// TIA Portal V21 export
// export: Created 2026-11-10T07:35:08.0372515Z, ExportSetting WithDefaults, DisplayName Totally Integrated Automation Portal, DisplayVersion V21 Update 3, DisplayName STEP 7 Professional, DisplayVersion V21 Update 3, DisplayName STEP 7 Safety, DisplayVersion V21, DisplayName Tech WebApplication, DisplayVersion V21, DisplayName WinCC Basic/Comfort/Advanced, DisplayVersion V21 Update 3, DisplayName WinCC Unified, DisplayVersion V21 Update 3
FUNCTION_BLOCK "FB_Lad_ex063"   // FB98, LAD
{ S7_Optimized_Access := 'TRUE' }
VERSION : 0.1
// stored: AutoNumber true, IsIECCheckEnabled false, IsRetainMemResEnabled false, MemoryReserve 100, SetENOAutomatically false, UDAEnableTagReadback false
   VAR_INPUT
      v_mode : Int;
      v_f_id : HW_SUBMODULE;
      v_code1 : Byte;
      v_code2 : Byte;
      v_len : UInt;
   END_VAR
   VAR_OUTPUT
      v_new : Bool;
      v_status : DWord;
      v_slot : HW_SUBMODULE;
      v_subslot : HW_SUBMODULE;
      v_index : UInt;
      v_rlen : UInt;
   END_VAR
   VAR_IN_OUT
      v_record : Array[0..99] of Byte;
   END_VAR
   VAR
      inst { S7_SetPoint := 'True'} : PRVREC;
   END_VAR
BEGIN

REGION Network 1: PRVREC - Make data record available
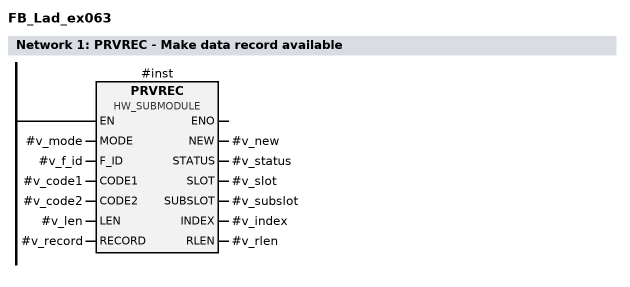
   RUNG wire#powerrail
      { S7_Templates := "[laddr_type := HW_SUBMODULE, ptr_type := Variant, len_type := UInt, id_type := HW_SUBMODULE]" } #inst.PRVREC(MODE := #v_mode, F_ID := #v_f_id, CODE1 := #v_code1, CODE2 := #v_code2, LEN := #v_len, NEW => #v_new, STATUS => #v_status, SLOT => #v_slot, SUBSLOT => #v_subslot, INDEX => #v_index, RLEN => #v_rlen, RECORD := #v_record)
   END_RUNG
   // the same network as SCL:
   #inst(MODE := #v_mode,   // PRVREC
         F_ID := #v_f_id,
         CODE1 := #v_code1,
         CODE2 := #v_code2,
         LEN := #v_len,
         RECORD := #v_record,
         NEW => #v_new,
         STATUS => #v_status,
         SLOT => #v_slot,
         SUBSLOT => #v_subslot,
         INDEX => #v_index,
         RLEN => #v_rlen);
END_REGION
END_FUNCTION_BLOCK
